(* IEC 61131-3 sources: STAR-PLC-Agent/results/raw/six_task_fullflow_20261114/PUB003/generation/sim_00, 1 file *)

(* ---- test_program.st ---- *)
PROGRAM PLC_PRG
VAR
 BenchStep : UDINT := 0;
 BenchCalls : UDINT := 0;
 BenchDone : BOOL := FALSE;
 BenchUut0 : FB_Task;
 BenchUut1 : FB_Task;
 TraceIn_Value : ARRAY[0..12] OF REAL;
 TraceIn_hiLevel : ARRAY[0..12] OF REAL;
 TraceIn_loLevel : ARRAY[0..12] OF REAL;
 TraceIn_hystWindow : ARRAY[0..12] OF REAL;
 TraceOut_hiAlarm : ARRAY[0..12] OF BOOL;
 TraceOut_loAlarm : ARRAY[0..12] OF BOOL;
 TraceOut_error : ARRAY[0..12] OF BOOL;
 TraceOut_status : ARRAY[0..12] OF WORD;
END_VAR

IF NOT BenchDone THEN
 CASE BenchStep OF
 0:
   BenchUut0.Value := REAL#50.0;
   BenchUut0.hiLevel := REAL#100.0;
   BenchUut0.loLevel := REAL#0.0;
   BenchUut0.hystWindow := REAL#10.0;
   TraceIn_Value[0] := BenchUut0.Value;
   TraceIn_hiLevel[0] := BenchUut0.hiLevel;
   TraceIn_loLevel[0] := BenchUut0.loLevel;
   TraceIn_hystWindow[0] := BenchUut0.hystWindow;
   BenchUut0();
   TraceOut_hiAlarm[0] := BenchUut0.hiAlarm;
   TraceOut_loAlarm[0] := BenchUut0.loAlarm;
   TraceOut_error[0] := BenchUut0.error;
   TraceOut_status[0] := BenchUut0.status;
   BenchCalls := BenchCalls + 1;
 1:
   BenchUut0.Value := REAL#110.0;
   BenchUut0.hiLevel := REAL#100.0;
   BenchUut0.loLevel := REAL#0.0;
   BenchUut0.hystWindow := REAL#10.0;
   TraceIn_Value[1] := BenchUut0.Value;
   TraceIn_hiLevel[1] := BenchUut0.hiLevel;
   TraceIn_loLevel[1] := BenchUut0.loLevel;
   TraceIn_hystWindow[1] := BenchUut0.hystWindow;
   BenchUut0();
   TraceOut_hiAlarm[1] := BenchUut0.hiAlarm;
   TraceOut_loAlarm[1] := BenchUut0.loAlarm;
   TraceOut_error[1] := BenchUut0.error;
   TraceOut_status[1] := BenchUut0.status;
   BenchCalls := BenchCalls + 1;
 2:
   BenchUut0.Value := REAL#95.0;
   BenchUut0.hiLevel := REAL#100.0;
   BenchUut0.loLevel := REAL#0.0;
   BenchUut0.hystWindow := REAL#10.0;
   TraceIn_Value[2] := BenchUut0.Value;
   TraceIn_hiLevel[2] := BenchUut0.hiLevel;
   TraceIn_loLevel[2] := BenchUut0.loLevel;
   TraceIn_hystWindow[2] := BenchUut0.hystWindow;
   BenchUut0();
   TraceOut_hiAlarm[2] := BenchUut0.hiAlarm;
   TraceOut_loAlarm[2] := BenchUut0.loAlarm;
   TraceOut_error[2] := BenchUut0.error;
   TraceOut_status[2] := BenchUut0.status;
   BenchCalls := BenchCalls + 1;
 3:
   BenchUut0.Value := REAL#85.0;
   BenchUut0.hiLevel := REAL#100.0;
   BenchUut0.loLevel := REAL#0.0;
   BenchUut0.hystWindow := REAL#10.0;
   TraceIn_Value[3] := BenchUut0.Value;
   TraceIn_hiLevel[3] := BenchUut0.hiLevel;
   TraceIn_loLevel[3] := BenchUut0.loLevel;
   TraceIn_hystWindow[3] := BenchUut0.hystWindow;
   BenchUut0();
   TraceOut_hiAlarm[3] := BenchUut0.hiAlarm;
   TraceOut_loAlarm[3] := BenchUut0.loAlarm;
   TraceOut_error[3] := BenchUut0.error;
   TraceOut_status[3] := BenchUut0.status;
   BenchCalls := BenchCalls + 1;
 4:
   BenchUut0.Value := REAL#-5.0;
   BenchUut0.hiLevel := REAL#100.0;
   BenchUut0.loLevel := REAL#0.0;
   BenchUut0.hystWindow := REAL#10.0;
   TraceIn_Value[4] := BenchUut0.Value;
   TraceIn_hiLevel[4] := BenchUut0.hiLevel;
   TraceIn_loLevel[4] := BenchUut0.loLevel;
   TraceIn_hystWindow[4] := BenchUut0.hystWindow;
   BenchUut0();
   TraceOut_hiAlarm[4] := BenchUut0.hiAlarm;
   TraceOut_loAlarm[4] := BenchUut0.loAlarm;
   TraceOut_error[4] := BenchUut0.error;
   TraceOut_status[4] := BenchUut0.status;
   BenchCalls := BenchCalls + 1;
 5:
   BenchUut0.Value := REAL#5.0;
   BenchUut0.hiLevel := REAL#100.0;
   BenchUut0.loLevel := REAL#0.0;
   BenchUut0.hystWindow := REAL#10.0;
   TraceIn_Value[5] := BenchUut0.Value;
   TraceIn_hiLevel[5] := BenchUut0.hiLevel;
   TraceIn_loLevel[5] := BenchUut0.loLevel;
   TraceIn_hystWindow[5] := BenchUut0.hystWindow;
   BenchUut0();
   TraceOut_hiAlarm[5] := BenchUut0.hiAlarm;
   TraceOut_loAlarm[5] := BenchUut0.loAlarm;
   TraceOut_error[5] := BenchUut0.error;
   TraceOut_status[5] := BenchUut0.status;
   BenchCalls := BenchCalls + 1;
 6:
   BenchUut0.Value := REAL#15.0;
   BenchUut0.hiLevel := REAL#100.0;
   BenchUut0.loLevel := REAL#0.0;
   BenchUut0.hystWindow := REAL#10.0;
   TraceIn_Value[6] := BenchUut0.Value;
   TraceIn_hiLevel[6] := BenchUut0.hiLevel;
   TraceIn_loLevel[6] := BenchUut0.loLevel;
   TraceIn_hystWindow[6] := BenchUut0.hystWindow;
   BenchUut0();
   TraceOut_hiAlarm[6] := BenchUut0.hiAlarm;
   TraceOut_loAlarm[6] := BenchUut0.loAlarm;
   TraceOut_error[6] := BenchUut0.error;
   TraceOut_status[6] := BenchUut0.status;
   BenchCalls := BenchCalls + 1;
 7:
   BenchUut1.Value := REAL#110.0;
   BenchUut1.hiLevel := REAL#100.0;
   BenchUut1.loLevel := REAL#0.0;
   BenchUut1.hystWindow := REAL#10.0;
   TraceIn_Value[7] := BenchUut1.Value;
   TraceIn_hiLevel[7] := BenchUut1.hiLevel;
   TraceIn_loLevel[7] := BenchUut1.loLevel;
   TraceIn_hystWindow[7] := BenchUut1.hystWindow;
   BenchUut1();
   TraceOut_hiAlarm[7] := BenchUut1.hiAlarm;
   TraceOut_loAlarm[7] := BenchUut1.loAlarm;
   TraceOut_error[7] := BenchUut1.error;
   TraceOut_status[7] := BenchUut1.status;
   BenchCalls := BenchCalls + 1;
 8:
   BenchUut1.Value := REAL#100.0;
   BenchUut1.hiLevel := REAL#100.0;
   BenchUut1.loLevel := REAL#0.0;
   BenchUut1.hystWindow := REAL#10.0;
   TraceIn_Value[8] := BenchUut1.Value;
   TraceIn_hiLevel[8] := BenchUut1.hiLevel;
   TraceIn_loLevel[8] := BenchUut1.loLevel;
   TraceIn_hystWindow[8] := BenchUut1.hystWindow;
   BenchUut1();
   TraceOut_hiAlarm[8] := BenchUut1.hiAlarm;
   TraceOut_loAlarm[8] := BenchUut1.loAlarm;
   TraceOut_error[8] := BenchUut1.error;
   TraceOut_status[8] := BenchUut1.status;
   BenchCalls := BenchCalls + 1;
 9:
   BenchUut1.Value := REAL#90.0;
   BenchUut1.hiLevel := REAL#100.0;
   BenchUut1.loLevel := REAL#0.0;
   BenchUut1.hystWindow := REAL#10.0;
   TraceIn_Value[9] := BenchUut1.Value;
   TraceIn_hiLevel[9] := BenchUut1.hiLevel;
   TraceIn_loLevel[9] := BenchUut1.loLevel;
   TraceIn_hystWindow[9] := BenchUut1.hystWindow;
   BenchUut1();
   TraceOut_hiAlarm[9] := BenchUut1.hiAlarm;
   TraceOut_loAlarm[9] := BenchUut1.loAlarm;
   TraceOut_error[9] := BenchUut1.error;
   TraceOut_status[9] := BenchUut1.status;
   BenchCalls := BenchCalls + 1;
 10:
   BenchUut1.Value := REAL#90.0;
   BenchUut1.hiLevel := REAL#100.0;
   BenchUut1.loLevel := REAL#100.0;
   BenchUut1.hystWindow := REAL#10.0;
   TraceIn_Value[10] := BenchUut1.Value;
   TraceIn_hiLevel[10] := BenchUut1.hiLevel;
   TraceIn_loLevel[10] := BenchUut1.loLevel;
   TraceIn_hystWindow[10] := BenchUut1.hystWindow;
   BenchUut1();
   TraceOut_hiAlarm[10] := BenchUut1.hiAlarm;
   TraceOut_loAlarm[10] := BenchUut1.loAlarm;
   TraceOut_error[10] := BenchUut1.error;
   TraceOut_status[10] := BenchUut1.status;
   BenchCalls := BenchCalls + 1;
 11:
   BenchUut1.Value := REAL#90.0;
   BenchUut1.hiLevel := REAL#100.0;
   BenchUut1.loLevel := REAL#0.0;
   BenchUut1.hystWindow := REAL#100.0;
   TraceIn_Value[11] := BenchUut1.Value;
   TraceIn_hiLevel[11] := BenchUut1.hiLevel;
   TraceIn_loLevel[11] := BenchUut1.loLevel;
   TraceIn_hystWindow[11] := BenchUut1.hystWindow;
   BenchUut1();
   TraceOut_hiAlarm[11] := BenchUut1.hiAlarm;
   TraceOut_loAlarm[11] := BenchUut1.loAlarm;
   TraceOut_error[11] := BenchUut1.error;
   TraceOut_status[11] := BenchUut1.status;
   BenchCalls := BenchCalls + 1;
 12:
   BenchUut1.Value := REAL#95.0;
   BenchUut1.hiLevel := REAL#100.0;
   BenchUut1.loLevel := REAL#0.0;
   BenchUut1.hystWindow := REAL#10.0;
   TraceIn_Value[12] := BenchUut1.Value;
   TraceIn_hiLevel[12] := BenchUut1.hiLevel;
   TraceIn_loLevel[12] := BenchUut1.loLevel;
   TraceIn_hystWindow[12] := BenchUut1.hystWindow;
   BenchUut1();
   TraceOut_hiAlarm[12] := BenchUut1.hiAlarm;
   TraceOut_loAlarm[12] := BenchUut1.loAlarm;
   TraceOut_error[12] := BenchUut1.error;
   TraceOut_status[12] := BenchUut1.status;
   BenchCalls := BenchCalls + 1;
 END_CASE;
 BenchStep := BenchStep + 1;
 IF BenchStep >= 13 THEN BenchDone := TRUE; END_IF;
END_IF;
END_PROGRAM
